(* IEC 61131-3 sources: codesys-framework/txt/application/WeVe Visu (library)/Controller/FB_NavBarController, 3 files *)

(* ---- HandleButtonClicks.method.st ---- *)
METHOD PRIVATE HandleButtonClicks : BOOL
VAR_INPUT
END_VAR

// --- BEGIN IMPLEMENTATION ---

IF _btnOperationalMode.RQ THEN
	SetFrame(iFrameToShow := 0);
END_IF

IF _btnSysParFR.RQ THEN
	SetFrame(iFrameToShow := 1);
END_IF

IF _btnSysParBuggy.RQ THEN
	SetFrame(iFrameToShow := 2);
END_IF

IF _btnJobManager.RQ THEN
	SetFrame(iFrameToShow := 3);
END_IF

IF _btnManualRequest.RQ THEN
	SetFrame(iFrameToShow := 4);
END_IF

IF _btnFeedRobot.RQ THEN
	SetFrame(iFrameToShow := 5);
END_IF

IF _btnYarnStorage.RQ THEN
	SetFrame(iFrameToShow := 6);
END_IF

IF _btnSysParSafety.RQ THEN
	SetFrame(iFrameToShow := 7);
END_IF

(* ---- ProcessFBs.method.st ---- *)
METHOD PRIVATE ProcessFBs : BOOL
VAR_INPUT
END_VAR

// --- BEGIN IMPLEMENTATION ---

_btnOperationalMode();
_btnParameters();
_btnSysParFR();
_btnSysParBuggy();
_btnSysParSafety();
_btnJobManager();
_btnManualRequest();
_btnFeedRobot();
_btnYarnStorage();

(* ---- SetFrame.method.st ---- *)
METHOD PRIVATE SetFrame : BOOL
VAR_INPUT
	iFrameToShow 		: UINT;
END_VAR

// --- BEGIN IMPLEMENTATION ---

iFrame := iFrameToShow;

xHideParameters := TRUE;
